// TwinCAT 3 PLC project Machine
// ProgramVersion: 3.1.4026.27
// libraries:
//   Tc2_Standard, * (Beckhoff Automation GmbH)
//   Tc2_System, * (Beckhoff Automation GmbH)
//   DemoLib,newest,Demo
// project tree:
//   DUTs/ E_FillStep.TcDUT, ST_DriveIn.TcDUT, ST_Recipe.TcDUT
//   GVLs/ GVL_IO.TcGVL, GVL_Parameters.TcGVL
//   / PlcTask.TcTTO
//   POUs/Equipment/ FB_Conveyor.TcPOU, FB_Sensor.TcPOU, FB_Valve.TcPOU
//   POUs/Experimental/ FB_Prototype.TcPOU
//   POUs/ MAIN.TcPOU, PRG_Lamp.TcPOU
//   POUs/Sequences/ FB_FillSequence.TcPOU
// real-time tasks:
//   TASK PlcTask: cycle T#10ms, priority 20, ADS port 350
// I/O:
//   DEVICE Device 1 (EtherCAT), AmsNetId 10.1.180.22.2.1
//     Term 1 (EK1100) [EK1100 EtherCAT Coupler (2A E-Bus)]
//       Term 2 (EL1008) [EL1008 8Ch. Dig. Input 24V, 3ms]
//       Term 3 (EL2008) [EL2008 8Ch. Dig. Output 24V, 0.5A]
//       Term 4 (EL3064) [EL3064 4Ch. Ana. Input 0-10V]
// variable links:
//   Machine/Machine Instance <-> Device 1 (EtherCAT)/Term 1 (EK1100)/Term 2 (EL1008)
//     PlcTask Inputs/GVL_IO.bStartButton <-> Channel 1/Input
//     PlcTask Inputs/GVL_IO.stDrive/bFault <-> Channel 4/Input
//     PlcTask Inputs/GVL_IO.stDrive/bReady <-> Channel 3/Input
//     PlcTask Inputs/MAIN.fbSensorLeft.bSignal <-> Channel 2/Input
//   Machine/Machine Instance <-> Device 1 (EtherCAT)/Term 1 (EK1100)/Term 3 (EL2008)
//     PlcTask Outputs/GVL_IO.aLamps[1] <-> Channel 3/Output
//     PlcTask Outputs/GVL_IO.aLamps[2] <-> Channel 4/Output
//     PlcTask Outputs/GVL_IO.bConveyorRun <-> Channel 2/Output
//     PlcTask Outputs/GVL_IO.bInletOpen <-> Channel 1/Output
//   Machine/Machine Instance <-> Device 1 (EtherCAT)/Term 1 (EK1100)/Term 4 (EL3064)
//     PlcTask Inputs/GVL_IO.nLevelRaw <-> AI Standard Channel 1/Value

CONFIGURATION Machine
    RESOURCE PLC ON TwinCAT3
        TASK PlcTask(INTERVAL := T#10ms, PRIORITY := 20);
        PROGRAM MAIN WITH PlcTask : MAIN;
    END_RESOURCE
END_CONFIGURATION

// ---- DUTs/E_FillStep.TcDUT
{attribute 'qualified_only'}
TYPE E_FillStep :
(
	Idle,
	OpenInlet,
	Filling,
	Settle,
	Done
) UINT;
END_TYPE

// ---- DUTs/ST_DriveIn.TcDUT
TYPE ST_DriveIn :
STRUCT
	bReady		: BOOL;
	bFault		: BOOL;
	nVelocity	: INT;
END_STRUCT
END_TYPE

// ---- DUTs/ST_Recipe.TcDUT
TYPE ST_Recipe :
STRUCT
	sName		: STRING(31);
	fTargetLevel	: T_Percent := 80;
	tSettle		: TIME := T#2S;
END_STRUCT
END_TYPE

// ---- GVLs/GVL_IO.TcGVL
VAR_GLOBAL
	bInletOpen		AT %Q*	: BOOL;
	bConveyorRun	AT %Q*	: BOOL;
	nLevelRaw		AT %I*	: INT;
	bStartButton	AT %I*	: BOOL;
	stDrive			AT %I*	: ST_DriveIn;
	aLamps			AT %Q*	: ARRAY[1..3] OF BOOL;
	bSpareOut		AT %Q*	: BOOL;	// spare: not linked
END_VAR

// ---- GVLs/GVL_Parameters.TcGVL
{attribute 'qualified_only'}
VAR_GLOBAL PERSISTENT
	stRecipe	: ST_Recipe := (sName := 'Default');
	fMaxSpeed	: LREAL := 1.5; // m/s
END_VAR

// ---- POUs/MAIN.TcPOU
PROGRAM MAIN
VAR
	fbInlet		: FB_Valve;
	fbConveyor	: FB_Conveyor;
	fbFill		: FB_FillSequence;
	uRaw		: U_Word;
	fbSensorLeft	: FB_Sensor;
	fbSensorRight	: FB_Sensor;
END_VAR

uRaw.nValue := INT_TO_WORD(GVL_IO.nLevelRaw);
fbFill(bStart := GVL_IO.bStartButton, fLevel := F_Clamp(WORD_TO_LREAL(uRaw.nValue) / 327.67, 0, 100), stRecipe := GVL_Parameters.stRecipe, iInlet := fbInlet);
fbInlet();
GVL_IO.bInletOpen := fbInlet.bOutput;

fbConveyor(bEnable := fbFill.bDone);
IF fbFill.bDone AND NOT fbConveyor.bRunning THEN
	fbConveyor.Speed := GVL_Parameters.fMaxSpeed;
	fbConveyor.Start();
END_IF
GVL_IO.bConveyorRun := fbConveyor.bRunning;
PRG_Lamp();

fbSensorLeft();
fbSensorRight();
GVL_IO.aLamps[1] := fbSensorLeft.bActive;
GVL_IO.aLamps[2] := fbSensorRight.bActive;
GVL_IO.aLamps[3] := GVL_IO.stDrive.bReady AND NOT GVL_IO.stDrive.bFault AND GVL_IO.stDrive.nVelocity > 0;

END_PROGRAM

// ---- POUs/Equipment/FB_Valve.TcPOU
FUNCTION_BLOCK FB_Valve EXTENDS FB_ValveBase
VAR_OUTPUT
	bOutput	: BOOL;
END_VAR

SUPER^();
bOutput := stStatus.eState = E_ValveState.Open OR stStatus.eState = E_ValveState.Opening;
IF stStatus.eState = E_ValveState.Opening THEN
	stStatus.eState := E_ValveState.Open;
ELSIF stStatus.eState = E_ValveState.Closing THEN
	stStatus.eState := E_ValveState.Closed;
END_IF

ACTION A_Reset:
stStatus.eState := E_ValveState.Closed;
stStatus.nCycles := 0;
bOutput := FALSE;
END_ACTION

METHOD Open : BOOL
VAR_INPUT
	bForce	: BOOL;
END_VAR
Open := SUPER^.Open(bForce := bForce);
IF Open THEN
	bOutput := TRUE;
END_IF
END_METHOD

END_FUNCTION_BLOCK

// ---- POUs/Equipment/FB_Conveyor.TcPOU
FUNCTION_BLOCK FB_Conveyor
VAR_INPUT
	bEnable	: BOOL;
END_VAR
VAR_OUTPUT
	bRunning	: BOOL;
END_VAR
VAR
	fSpeed		: LREAL;
	bStartReq	: BOOL;
END_VAR

bRunning := bEnable AND bStartReq AND fSpeed > 0;

PROPERTY Speed : LREAL
GET // PUBLIC
Speed := fSpeed;
END_GET
SET // PUBLIC
fSpeed := F_Clamp(Speed, 0, GVL_Parameters.fMaxSpeed);
END_SET
END_PROPERTY

METHOD Start : BOOL
bStartReq := bEnable;
Start := bStartReq;
END_METHOD

METHOD Stop
bStartReq := FALSE;
END_METHOD

END_FUNCTION_BLOCK

// ---- POUs/Sequences/FB_FillSequence.TcPOU
FUNCTION_BLOCK FB_FillSequence
VAR_INPUT
	bStart		: BOOL;
	fLevel		: T_Percent;
	stRecipe	: ST_Recipe;
	iInlet		: I_Valve;
END_VAR
VAR_OUTPUT
	eStep		: E_FillStep;
	bDone		: BOOL;
END_VAR
VAR
	tonSettle	: TON;
END_VAR

CASE eStep OF
	E_FillStep.Idle:
		bDone := FALSE;
		IF bStart THEN
			eStep := E_FillStep.OpenInlet;
		END_IF

	E_FillStep.OpenInlet:
		IF iInlet.Open(bForce := FALSE) THEN
			eStep := E_FillStep.Filling;
		END_IF

	E_FillStep.Filling:
		IF fLevel >= stRecipe.fTargetLevel THEN
			iInlet.Close();
			eStep := E_FillStep.Settle;
		END_IF

	E_FillStep.Settle:
		tonSettle(IN := TRUE, PT := stRecipe.tSettle);
		IF tonSettle.Q THEN
			tonSettle(IN := FALSE);
			eStep := E_FillStep.Done;
		END_IF

	E_FillStep.Done:
		bDone := TRUE;
		IF NOT bStart THEN
			eStep := E_FillStep.Idle;
		END_IF
END_CASE

END_FUNCTION_BLOCK

// ---- POUs/Equipment/FB_Sensor.TcPOU
FUNCTION_BLOCK FB_Sensor
VAR_OUTPUT
	bActive	: BOOL;
END_VAR
VAR
	bSignal	AT %I*	: BOOL;
END_VAR

bActive := bSignal;

END_FUNCTION_BLOCK

// ---- POUs/PRG_Lamp.TcPOU
PROGRAM PRG_Lamp
VAR
	bLamp	: BOOL;
END_VAR

END_PROGRAM

// ---- POUs/Experimental/FB_Prototype.TcPOU
FUNCTION_BLOCK FB_Prototype
VAR
	nCount	: INT;
END_VAR

nCount := nCount + UnknownSymbol; // not built: the folder is excluded from the build

END_FUNCTION_BLOCK
